Fanuc KAREL source: KB00164.KL

PROGRAM KB00164
%NOLOCKGROUP
%ENVIRONMENT FLBT
VAR
  P1: FILE
  P2: INTEGER
  P3: INTEGER
BEGIN
  P2 = 1
  P3 = 1
  SET_FILE_POS(P1, P2, P3)
END KB00164
